// TIA Portal V21 export
// export: Created 2026-11-10T19:16:29.8458396Z, ExportSetting WithDefaults, DisplayName Totally Integrated Automation Portal, DisplayVersion V21 Update 3, DisplayName STEP 7 Professional, DisplayVersion V21 Update 3, DisplayName STEP 7 Safety, DisplayVersion V21, DisplayName Tech WebApplication, DisplayVersion V21, DisplayName WinCC Basic/Comfort/Advanced, DisplayVersion V21 Update 3, DisplayName WinCC Unified, DisplayVersion V21 Update 3
DATA_BLOCK "DB_12Std"   // DB2
{ S7_Optimized_Access := 'FALSE' }
VERSION : 0.1
// stored: AutoNumber true, DBAccessibleFromOPCUA true, IsOnlyStoredInLoadMemory false, IsWriteProtectedInAS false
   VAR
      b0 : Bool;
      w : Word;
      i : Int := -4;
      r : Real;
      s : String[6];
      arr : Array[0..3] of Int;
      u { S7_SetPoint := 'True'} : "UDT_12";
   END_VAR
BEGIN
   arr[2] := 22;
END_DATA_BLOCK
